FUNCTION_BLOCK PUBLIC FB_Dissolving EXTENDS FB_SFC_Cycle IMPLEMENTS ITF_FB_SFC_Cycle
VAR_INPUT
END_VAR
VAR_OUTPUT
END_VAR
VAR
	step: INT;
	i: INT;
	ton_Blending_Speed: TON;
	tBlending: TIME;
	tBlending_count: TIME;
	ptTemp: DINT;
	tBlendingRemainTime: DINT;
	realTemp: REAL;
	fBlendingPercenatge: DINT;
END_VAR

VAR_IN_OUT
	fb_TriBlender			: FB_Pump;
END_VAR

m_Set_SFCFlags_Reference();
act_Oper();
IF g_HMI_Panel.stPLC_To_VisuPLC.iActual_Component<>0 THEN
	ptTemp:=TIME_TO_DINT(g_HMI_Panel.stPLC_To_VisuPLC.arr_Component[g_HMI_Panel.stPLC_To_VisuPLC.iActual_Component].tBlendingDuration);
ELSE;
	ptTemp:=0;
END_IF

tBlendingRemainTime:=ptTemp - TIME_TO_DINT(tBlending);
IF ptTemp<>0 THEN;
	realTemp:=(DINT_TO_REAL(tBlendingRemainTime)/DINT_TO_REAL(ptTemp)*100.0);
	fBlendingPercenatge:=TRUNC(realTemp);
END_IF

ACTION _aChek_if_Done_active:
bStepDone:=FALSE;
IF g_HMI_Panel.stPLC_To_VisuPLC.iActual_Component >= 10 THEN;
	bStepDone:=TRUE;
END_IF
END_ACTION

ACTION _aComponent_Blending_active:
bStepDone:=FALSE;
IF tBlending > g_HMI_Panel.stPLC_To_VisuPLC.arr_Component[g_HMI_Panel.stPLC_To_VisuPLC.iActual_Component].tBlendingDuration THEN;
	bStepDone:=TRUE;
	g_HMI_Panel.stPLC_To_VisuPLC.bBlending_Active:=FALSE;
END_IF

fb_TriBlender.m_Run(RPM:=g_HMI_Panel.stPLC_To_VisuPLC.arr_Component[g_HMI_Panel.stPLC_To_VisuPLC.iActual_Component].rFlowRate_Blending);

ton_Blending_Speed(PT:=T#2S);
IF TRUE 
AND fb_TriBlender.m_Get_Speed() >= g_HMI_Panel.stPLC_To_VisuPLC.arr_Component[g_HMI_Panel.stPLC_To_VisuPLC.iActual_Component].rFlowRate_Blending - 10
AND fb_TriBlender.m_Get_Speed() <= g_HMI_Panel.stPLC_To_VisuPLC.arr_Component[g_HMI_Panel.stPLC_To_VisuPLC.iActual_Component].rFlowRate_Blending + 10
THEN;
	ton_Blending_Speed.IN:=TRUE;
ELSE;
	ton_Blending_Speed.IN:=FALSE;
END_IF

IF ton_Blending_Speed.Q THEN;
	tBlending:=tBlending + T#10MS; // scan Time
ELSE;
	
END_IF
END_ACTION

ACTION _aComponent_Blending_entry:
g_HMI_Panel.stPLC_To_VisuPLC.bDissolving_Active:=FALSE;
g_HMI_Panel.stPLC_To_VisuPLC.bBlending_Active:=TRUE;
END_ACTION

ACTION _aDissolving_Done_entry:
bDisolvingProcess_Done:=TRUE;
END_ACTION

ACTION _aInit_Dissolve_exit:
step:=0;
g_HMI_Panel.stPLC_To_VisuPLC.iActual_Component:=0;
g_HMI_Panel.stPLC_To_VisuPLC.bDissolving_Active:=FALSE;
g_HMI_Panel.stPLC_To_VisuPLC.bBlending_Active:=FALSE;
bRun:=FALSE;
END_ACTION

ACTION _aReady_exit:
g_HMI_Panel.stPLC_To_VisuPLC.iActual_Component:=1;
g_HMI_Panel.stPLC_To_VisuPLC.bDissolving_Active:=FALSE;
END_ACTION

ACTION _arepeat_stage_active:
bStepDone:=NOT g_HMI_Panel.stVisuPLC_To_PLC.bActualComponentDisolving_Done;
END_ACTION

ACTION _aSet_Next_Component_active:
bStepDone:=FALSE;
IF g_HMI_Panel.stVisuPLC_To_PLC.bActualComponentDisolving_Done THEN;
	bStepDone:=TRUE;
END_IF

IF g_HMI_Panel.stVisuPLC_To_PLC.bPauseTriBlender THEN;
	fb_TriBlender.m_Stop();
ELSE;
	fb_TriBlender.m_Run(RPM:=g_HMI_Panel.stVisuPLC_To_PLC.RPM_setPoint);
END_IF
END_ACTION

ACTION _aSet_Next_Component_entry:
g_HMI_Panel.stPLC_To_VisuPLC.bDissolving_Active:=FALSE;
g_HMI_Panel.stPLC_To_VisuPLC.bBlending_Active:=FALSE;
g_HMI_Panel.stPLC_To_VisuPLC.iActual_Component:=g_HMI_Panel.stPLC_To_VisuPLC.iActual_Component+1;

FOR i:=g_HMI_Panel.stPLC_To_VisuPLC.iActual_Component TO 10 DO
	IF g_HMI_Panel.stPLC_To_VisuPLC.arr_Component[i].rWeight>0 THEN;
		g_HMI_Panel.stPLC_To_VisuPLC.iActual_Component:=i;
		g_HMI_Panel.stPLC_To_VisuPLC.bDissolving_Active:=TRUE;
		EXIT;
	END_IF
END_FOR

tBlending:=T#0S;
END_ACTION

ACTION act_Oper:
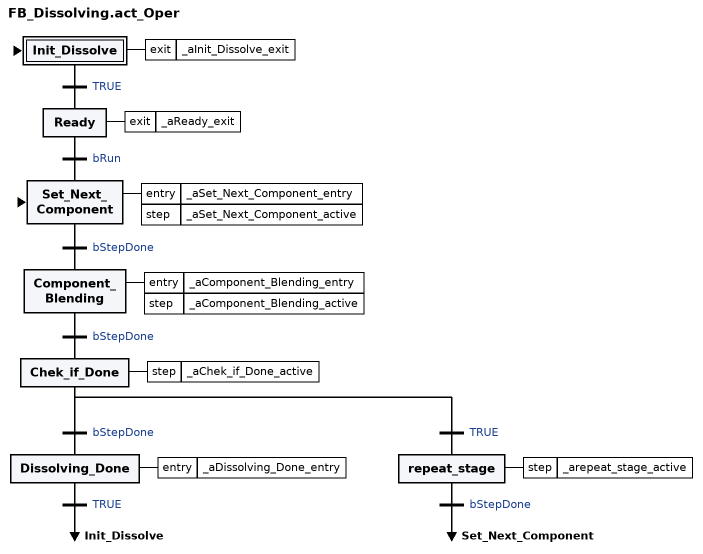
INITIAL_STEP Init_Dissolve:
    _aInit_Dissolve_exit(P0);  // exit action
END_STEP
TRANSITION FROM Init_Dissolve TO Ready
    := TRUE;
END_TRANSITION
STEP Ready:
    _aReady_exit(P0);  // exit action
END_STEP
TRANSITION FROM Ready TO Set_Next_Component
    := bRun;
END_TRANSITION
STEP Set_Next_Component:
    _aSet_Next_Component_entry(P1);  // entry action
    _aSet_Next_Component_active(N);  // step action
END_STEP
TRANSITION FROM Set_Next_Component TO Component_Blending
    := bStepDone;
END_TRANSITION
STEP Component_Blending:
    _aComponent_Blending_entry(P1);  // entry action
    _aComponent_Blending_active(N);  // step action
END_STEP
TRANSITION FROM Component_Blending TO Chek_if_Done
    := bStepDone;
END_TRANSITION
STEP Chek_if_Done:
    _aChek_if_Done_active(N);  // step action
END_STEP
TRANSITION FROM Chek_if_Done TO Dissolving_Done
    := bStepDone;
END_TRANSITION
TRANSITION FROM Chek_if_Done TO repeat_stage
    := TRUE;
END_TRANSITION
STEP repeat_stage:
    _arepeat_stage_active(N);  // step action
END_STEP
TRANSITION FROM repeat_stage TO Set_Next_Component
    := bStepDone;
END_TRANSITION
STEP Dissolving_Done:
    _aDissolving_Done_entry(P1);  // entry action
END_STEP
TRANSITION FROM Dissolving_Done TO Init_Dissolve
    := TRUE;
END_TRANSITION
// branch label Branch0_act_Oper
END_ACTION

METHOD m_Set_SFCFlags_Reference : BOOL
//Set reference to SFC flags

refSFC.SFCInit REF= SFCInit;
refSFC.SFCReset REF= SFCReset;
refSFC.SFCError REF= SFCError;
refSFC.SFCEnableLimit REF= SFCEnableLimit;
refSFC.SFCErrorStep REF= SFCErrorStep;
refSFC.SFCErrorPOU REF= SFCErrorPOU;
refSFC.SFCQuitError REF= SFCQuitError;
refSFC.SFCPause REF= SFCPause;
refSFC.SFCTrans REF= SFCTrans;
refSFC.SFCCurrentStep REF= SFCCurrentStep;
refSFC.SFCTip REF= SFCTip;
refSFC.SFCTipMode REF= SFCTipMode;

// Cycle handle for SFC
m_SFC_Handle();
END_METHOD

END_FUNCTION_BLOCK

(* stored: Version 1.1.0.1, ProductVersion 3.1.4024.15
   POU FB_Dissolving: Id {61fb2bea-f425-42ba-8eea-35efb6847cdf}, SpecialFunc None
   Action _aChek_if_Done_active: Id {28a6cd2f-fcb4-4026-979e-d8afebb2d7fb}
   Action _aComponent_Blending_active: Id {49c635d9-8cb2-43c9-af22-31b599cbdffb}
   Action _aComponent_Blending_entry: Id {4c0e6d76-310b-4245-93e0-c7c557bef00e}
   Action _aDissolving_Done_entry: Id {fb0791ee-288b-493f-9dec-4045da4634b4}
   Action _aInit_Dissolve_exit: Id {d2eef2f7-7f78-404f-8147-d7c62309e56f}
   Action _aReady_exit: Id {9fefdedd-c232-4791-9377-8e14ef06db2d}
   Action _arepeat_stage_active: Id {74b73a03-d912-4c2f-a00f-2441cd673961}
   Action _aSet_Next_Component_active: Id {bdf66cc9-1360-4ca9-a4b1-8e42f5ad1b30}
   Action _aSet_Next_Component_entry: Id {0b708c24-9fee-4a9b-ba4f-f7202d8afeaa}
   Action act_Oper: Id {1fc2d52a-af85-41c6-9e56-9caeb95a124c}
   Method m_Set_SFCFlags_Reference: Id {81b13ccf-b7e9-484f-a8de-970add58bd6f} *)
